// TIA Portal V21 export
// export: Created 2026-11-07T15:50:50.6268125Z, ExportSetting WithDefaults, DisplayName Totally Integrated Automation Portal, DisplayVersion V21, DisplayName STEP 7 Professional, DisplayVersion V21, DisplayName STEP 7 Safety, DisplayVersion V21, DisplayName Tech WebApplication, DisplayVersion V21, DisplayName WinCC Basic/Comfort/Advanced, DisplayVersion V21, DisplayName WinCC Unified, DisplayVersion V21
Screen "R06a_MoveH"  1024x768, Number=45, Template=Tpl
  ScreenLayer 
    IOField "P_CraneX" at 10,10 size 100x30  DataFormat=Decimal, FormatPattern=999.999, Mode=Output, StyleItem=I/O field
      HorizontalMovementAnimation "HorizontalMovementAnimation"  RangeEnd=100, XDelta=200, XPosEnd=210
        tag 
      ProcessValue := P_Cell
